DATA_BLOCK "naut_SfcSimDivConv_DB"
{ S7_Optimized_Access := 'TRUE' }
VERSION : 0.1
"naut_SfcSimDivConv"

BEGIN

END_DATA_BLOCK
